TYPE ST_SwitchControlData :
STRUCT
    bShortClick      : BOOL;
    nShortClickCount : USINT;
    bLongClick       : BOOL;
    bIsHeld          : BOOL;
    bHoldReleased    : BOOL;
END_STRUCT
END_TYPE

(* stored: Version 1.1.0.1, ProductVersion 3.1.4026.20
   DUT ST_SwitchControlData: Id {A9E21D47-5C83-4B10-9F62-1D7A3C8E5001} *)
